RoboDK station: PRBE_Operateur_v2.rdk

Station PRBE_Operateur_v2 (saved by RoboDK 6.0.4). Poses are relative to the parent item; angles as X-Y-Z fixed-axis rotations.
  - object Manikin_1 at (0, 0, 0) mm, geometry from Manikin_1.STEP
  - frame Human_Base at (0, 958, 0) mm
    - item type 7 Manikin_1-bassin
    - item type 7 Manikin_1-torso
    - item type 7 Manikin_1-tete
    - frame hipL_abduction at (63.26, -78.51, -37.42) mm
      - frame hipL_flexion at (0, 0, 0) mm
        - frame hipL_rotation at (0, 0, 0) mm
          - item type 7 Manikin_1-cuisse_g
          - frame kneeL_flexion at (67.44, -393.44, -12.97) mm
            - item type 7 Manikin_1-tibia_g
            - frame ankleL_flexion at (42.46, -394.54, 0) mm
              - item type 7 Manikin_1-pied_g
    - frame shoulderL_abduction at (206.4, 423.68, 12.96) mm, rotated rx 0 ry 0 rz -42 deg
      - frame shoulderL_flexion at (0, 0, 0) mm
        - frame shoulderL_rotation at (0, 0, 0) mm
          - item type 7 Manikin_1-bras_g
          - frame elbowL_flexion at (155.8, -191.9, 27.9) mm
            - item type 7 Manikin_1-avant_bras_g
            - frame wristL_flexion at (148.7, -146.81, 80.89) mm
              - frame wristL_deviation at (0, 0, 0) mm
                - item type 7 Manikin_1-main_g
    - frame hipR_abduction at (-70.11, -75.34, -37.06) mm
      - frame hipR_flexion at (0, 0, 0) mm
        - frame hipR_rotation at (0, 0, 0) mm
          - item type 7 Manikin_1-cuisse_d
          - frame kneeR_flexion at (-86.5, -385.51, -37.91) mm
            - item type 7 Manikin_1-tibia_d_1
            - item type 7 Manikin_1-tibia_d_2
            - frame ankleR_flexion at (-60.5, -382.31, -26.03) mm
              - item type 7 Manikin_1-pied_d_1
              - item type 7 Manikin_1-pied_d_2
    - frame shoulderR_abduction at (-133.98, 420.49, -26.02) mm
      - frame shoulderR_flexion at (0, 0, 0) mm
        - frame shoulderR_rotation at (0, 0, 0) mm
          - item type 7 Manikin_1-bras_d
          - frame elbowR_flexion at (-80.76, -228.86, 52.14) mm
            - item type 7 Manikin_1-avant_bras_d
            - frame wristR_flexion at (-76.34, -195.54, 87.27) mm
              - frame wristR_deviation at (0, 0, 0) mm
                - item type 7 Manikin_1-main_d
  - Python program Mouvement_v2 (listed below)
  - Python program Marche_Militaire (listed below)
  - Python program Marche_Avant (listed below)

--- Python program Mouvement_v2 ---
# -*- coding: utf-8 -*-
"""
Mouvement_v2.py — MODELE pour piloter l'operateur v2 (22 DDL).

A LANCER DANS ROBODK (clic droit > Run) depuis la station PRBE_Operateur_v2,
operateur en pose NEUTRE (le script capture le repos au demarrage).

PRINCIPE :
  - chaque DDL = un repere nomme (ex: "hipR_flexion") qui tourne sur UN axe.
  - bouge("nom_du_ddl", angle_en_degres) tourne ce DDL depuis le repos.
  - les angles sont automatiquement borns aux limites du corps humain.
"""
from robolink import Robolink
from robodk.robomath import rotx, roty, rotz
import math
import time

RDK = Robolink()

# ---- Les 22 DDL : nom -> (axe, limite_basse_deg, limite_haute_deg) ----
DDL = {
    # JAMBE DROITE (5)
    "hipR_abduction": ("z", -45, 30),   "hipR_flexion": ("x", -120, 15),  "hipR_rotation": ("y", -45, 45),
    "kneeR_flexion":  ("x", 0, 135),    "ankleR_flexion": ("x", -30, 50),
    # JAMBE GAUCHE (5)
    "hipL_abduction": ("z", -30, 45),   "hipL_flexion": ("x", -120, 15),  "hipL_rotation": ("y", -45, 45),
    "kneeL_flexion":  ("x", 0, 135),    "ankleL_flexion": ("x", -30, 50),
    # BRAS DROIT (6)
    "shoulderR_abduction": ("z", -135, 90), "shoulderR_flexion": ("x", -90, 90), "shoulderR_rotation": ("y", -45, 180),
    "elbowR_flexion": ("x", 0, 145),
    "wristR_flexion": ("x", -50, 60),   "wristR_deviation": ("z", -30, 20),
    # BRAS GAUCHE (6)
    "shoulderL_abduction": ("z", -90, 135), "shoulderL_flexion": ("x", -90, 90), "shoulderL_rotation": ("y", -45, 180),
    "elbowL_flexion": ("x", 0, 145),
    "wristL_flexion": ("x", -50, 60),   "wristL_deviation": ("z", -30, 20),
}

ROT = {"x": rotx, "y": roty, "z": rotz}
F = {nom: RDK.Item(nom) for nom in DDL}            # les reperes
REST = {nom: F[nom].Pose() for nom in DDL}         # pose neutre (capturee au demarrage)


def bouge(nom, deg):
    """Tourne un DDL de `deg` degres depuis le repos (born aux limites)."""
    axe, lo, hi = DDL[nom]
    deg = max(lo, min(hi, deg))                    # ne depasse pas le corps humain
    F[nom].setPose(REST[nom] * ROT[axe](math.radians(deg)))


def neutre():
    """Remet tout l'operateur droit."""
    for nom in DDL:
        F[nom].setPose(REST[nom])


# =======================================================================
# TON CODE ICI. Exemples :
# =======================================================================

# --- EXEMPLE 1 : une pose (lever le bras droit + plier le coude) ---
bouge("shoulderR_flexion", -70)   # bras droit vers l'avant
bouge("elbowR_flexion", 90)       # coude plie
RDK.Render(True)
time.sleep(1)

# --- EXEMPLE 2 : une petite animation (le bras qui salue) ---
neutre()
bouge("shoulderR_abduction", 80)  # bras leve sur le cote
for i in range(6):
    RDK.Render(False)
    bouge("elbowR_flexion", 30 + 40 * (i % 2))   # avant-bras qui va et vient
    RDK.Render(True)
    time.sleep(0.3)

neutre()
RDK.Render(True)
print("Fini.")

--- Python program Marche_Militaire ---
# -*- coding: utf-8 -*-
"""
Marche_Militaire.py — L'operateur marque le pas (marche militaire sur place).

A LANCER DANS ROBODK (clic droit > Run) depuis la station avec le rig 22 DDL,
operateur en pose NEUTRE (le script capture le repos au demarrage).

Principe de la marche militaire :
  - genoux qui montent haut, alternes
  - bras RAIDES (coude quasi tendu) qui balancent en OPPOSITION des jambes
  - buste droit (il est fige, parfait pour un militaire)

Regle les amplitudes/vitesse dans la section REGLAGES.
"""
from robolink import Robolink
from robodk.robomath import rotx, roty, rotz
import math
import time

RDK = Robolink()

# ---- Les 22 DDL : nom -> (axe, limite_basse_deg, limite_haute_deg) ----
DDL = {
    # JAMBE DROITE (5)
    "hipR_abduction": ("z", -45, 30),   "hipR_flexion": ("x", -120, 15),  "hipR_rotation": ("y", -45, 45),
    "kneeR_flexion":  ("x", 0, 135),    "ankleR_flexion": ("x", -30, 50),
    # JAMBE GAUCHE (5)
    "hipL_abduction": ("z", -30, 45),   "hipL_flexion": ("x", -120, 15),  "hipL_rotation": ("y", -45, 45),
    "kneeL_flexion":  ("x", 0, 135),    "ankleL_flexion": ("x", -30, 50),
    # BRAS DROIT (6)
    "shoulderR_abduction": ("z", -135, 90), "shoulderR_flexion": ("x", -90, 90), "shoulderR_rotation": ("y", -45, 180),
    "elbowR_flexion": ("x", 0, 145),
    "wristR_flexion": ("x", -50, 60),   "wristR_deviation": ("z", -30, 20),
    # BRAS GAUCHE (6)
    "shoulderL_abduction": ("z", -90, 135), "shoulderL_flexion": ("x", -90, 90), "shoulderL_rotation": ("y", -45, 180),
    "elbowL_flexion": ("x", 0, 145),
    "wristL_flexion": ("x", -50, 60),   "wristL_deviation": ("z", -30, 20),
}

ROT = {"x": rotx, "y": roty, "z": rotz}
F = {nom: RDK.Item(nom) for nom in DDL}            # les reperes
REST = {nom: F[nom].Pose() for nom in DDL}         # pose neutre (capturee au demarrage)


def bouge(nom, deg):
    """Tourne un DDL de `deg` degres depuis le repos (borne aux limites)."""
    axe, lo, hi = DDL[nom]
    deg = max(lo, min(hi, deg))
    F[nom].setPose(REST[nom] * ROT[axe](math.radians(deg)))


def neutre():
    """Remet tout l'operateur droit."""
    for nom in DDL:
        F[nom].setPose(REST[nom])


# =======================================================================
# REGLAGES de la marche militaire
# =======================================================================
HANCHE = 55      # levee de cuisse (deg) — genou haut
GENOU = 65       # pliage du genou quand la jambe monte (deg)
CHEVILLE = 15    # pointe de pied quand la jambe est levee (deg)
BRAS_AV = -45    # bras vers l'AVANT (deg, negatif = devant)
BRAS_ARR = 20    # bras vers l'ARRIERE (deg)
COUDE = 8        # coude quasi tendu = bras raide militaire
NB_PAS = 8       # nombre de pas au total
IMAGES_PAR_PAS = 12   # fluidite (images par pas)
DT = 0.04        # pause entre images (s) — plus petit = plus rapide


def pose_marche(ph):
    """Pose complete de la marche pour une phase `ph` (radians).
       Jambe droite levee sur [0, pi], jambe gauche sur [pi, 2pi]."""
    s = math.sin(ph)
    lift_d = max(0.0, s)     # jambe droite qui monte
    lift_g = max(0.0, -s)    # jambe gauche qui monte

    # jambes : genou haut + pointe de pied
    bouge("hipR_flexion", -HANCHE * lift_d)
    bouge("kneeR_flexion", GENOU * lift_d)
    bouge("ankleR_flexion", CHEVILLE * lift_d)
    bouge("hipL_flexion", -HANCHE * lift_g)
    bouge("kneeL_flexion", GENOU * lift_g)
    bouge("ankleL_flexion", CHEVILLE * lift_g)

    # bras raides, en opposition : bras droit devant quand jambe gauche monte
    u_d = (1.0 - s) / 2.0    # 0 = bras D derriere, 1 = bras D devant
    u_g = (1.0 + s) / 2.0
    bouge("shoulderR_flexion", BRAS_ARR + (BRAS_AV - BRAS_ARR) * u_d)
    bouge("shoulderL_flexion", BRAS_ARR + (BRAS_AV - BRAS_ARR) * u_g)
    bouge("elbowR_flexion", COUDE)
    bouge("elbowL_flexion", COUDE)


def marche(nb_pas=NB_PAS, images_par_pas=IMAGES_PAR_PAS, dt=DT):
    """Anime la marche militaire sur place."""
    for i in range(nb_pas * images_par_pas + 1):
        ph = math.pi * i / images_par_pas      # 1 pas = une demi-periode
        RDK.Render(False)
        pose_marche(ph)
        RDK.Render(True)
        time.sleep(dt)
    neutre()
    RDK.Render(True)


if __name__ == "__main__":
    print("Marche militaire : {} pas...".format(NB_PAS))
    marche()
    print("Repos !")

--- Python program Marche_Avant ---
# -*- coding: utf-8 -*-
"""
Marche_Avant.py — L'operateur marche TOUT DROIT devant lui (marche naturelle).

A LANCER DANS ROBODK (clic droit > Run) depuis la station avec le rig 22 DDL,
operateur au repos / garde-a-vous (le script capture le repos au demarrage).

Principe :
  - hanches qui balancent avant/arriere, genou qui se plie pendant le balance
  - bras souples en opposition des jambes (coude legerement plie)
  - le CORPS AVANCE a la vitesse des pas (longueur de pas calculee depuis
    l'amplitude de hanche) -> pas de glisse visible
  - il marche vers SON regard (+Z monde). A la fin, il REVIENT au centre
    (position d'origine de Human_Base).

Regle les amplitudes/vitesse dans la section REGLAGES.
"""
from robolink import Robolink
from robodk.robomath import rotx, roty, rotz, transl
import math
import time

RDK = Robolink()

# ---- Les 22 DDL : nom -> (axe, limite_basse_deg, limite_haute_deg) ----
DDL = {
    # JAMBE DROITE (5)
    "hipR_abduction": ("z", -45, 30),   "hipR_flexion": ("x", -120, 15),  "hipR_rotation": ("y", -45, 45),
    "kneeR_flexion":  ("x", 0, 135),    "ankleR_flexion": ("x", -30, 50),
    # JAMBE GAUCHE (5)
    "hipL_abduction": ("z", -30, 45),   "hipL_flexion": ("x", -120, 15),  "hipL_rotation": ("y", -45, 45),
    "kneeL_flexion":  ("x", 0, 135),    "ankleL_flexion": ("x", -30, 50),
    # BRAS DROIT (6)
    "shoulderR_abduction": ("z", -135, 90), "shoulderR_flexion": ("x", -90, 90), "shoulderR_rotation": ("y", -45, 180),
    "elbowR_flexion": ("x", 0, 145),
    "wristR_flexion": ("x", -50, 60),   "wristR_deviation": ("z", -30, 20),
    # BRAS GAUCHE (6)
    "shoulderL_abduction": ("z", -90, 135), "shoulderL_flexion": ("x", -90, 90), "shoulderL_rotation": ("y", -45, 180),
    "elbowL_flexion": ("x", 0, 145),
    "wristL_flexion": ("x", -50, 60),   "wristL_deviation": ("z", -30, 20),
}

ROT = {"x": rotx, "y": roty, "z": rotz}
F = {nom: RDK.Item(nom) for nom in DDL}            # les reperes
REST = {nom: F[nom].Pose() for nom in DDL}         # pose de repos (capturee au demarrage)
BASE = RDK.Item("Human_Base")
BASE_REST = BASE.Pose()                            # position de depart du corps
HOME = transl(0, 958, 0)                           # position d'origine (au centre, 1er repere)


def bouge(nom, deg):
    """Tourne un DDL de `deg` degres depuis le repos (borne aux limites)."""
    axe, lo, hi = DDL[nom]
    deg = max(lo, min(hi, deg))
    F[nom].setPose(REST[nom] * ROT[axe](math.radians(deg)))


def neutre():
    """Remet les articulations au repos (le corps reste ou il est)."""
    for nom in DDL:
        F[nom].setPose(REST[nom])


# =======================================================================
# REGLAGES de la marche
# =======================================================================
HANCHE_AV = 30    # jambe vers l'avant (deg)
HANCHE_ARR = 12   # jambe vers l'arriere (deg)
GENOU = 50        # pliage du genou pendant le balance (deg)
CHEVILLE = 8      # pointe de pied relevee pendant le balance (deg)
BRAS_AV = 25      # bras vers l'avant (deg)
BRAS_ARR = 15     # bras vers l'arriere (deg)
COUDE = 20        # coude legerement plie (marche naturelle)
NB_PAS = 8        # nombre de pas
IMAGES_PAR_PAS = 14   # fluidite
DT = 0.04         # pause entre images (s)

LONGUEUR_JAMBE = 790.0   # hanche -> cheville (mm, mesure sur le modele)
SENS = +1                # +1 = devant lui (+Z monde). Mets -1 pour marche arriere.

# longueur d'un pas deduite du balancement de hanche (pour avancer sans glisser)
LONGUEUR_PAS = LONGUEUR_JAMBE * (math.sin(math.radians(HANCHE_AV)) + math.sin(math.radians(HANCHE_ARR)))


def pose_pas(ph):
    """Pose de marche pour une phase `ph` (radians). Jambe droite devant sur [0, pi]."""
    s = math.sin(ph)
    # hanches : avant = negatif (amplitude asymetrique avant/arriere)
    a = (HANCHE_AV + HANCHE_ARR) / 2.0
    c = (HANCHE_AV - HANCHE_ARR) / 2.0
    bouge("hipR_flexion", -(a * s + c))
    bouge("hipL_flexion", -(a * -s + c))
    # genou plie pendant le balance (jambe qui revient vers l'avant)
    bouge("kneeR_flexion", GENOU * max(0.0, math.cos(ph)))
    bouge("kneeL_flexion", GENOU * max(0.0, -math.cos(ph)))
    # pointe de pied relevee pendant le balance (pour ne pas racler le sol)
    bouge("ankleR_flexion", -CHEVILLE * max(0.0, math.cos(ph)))
    bouge("ankleL_flexion", -CHEVILLE * max(0.0, -math.cos(ph)))
    # bras en opposition, coude souple
    sa = (BRAS_AV + BRAS_ARR) / 2.0
    sc = (BRAS_ARR - BRAS_AV) / 2.0
    bouge("shoulderR_flexion", sa * s + sc)
    bouge("shoulderL_flexion", -sa * s + sc)
    bouge("elbowR_flexion", COUDE)
    bouge("elbowL_flexion", COUDE)


def avance(dist):
    """Place le corps a `dist` mm devant sa position de depart."""
    BASE.setPose(BASE_REST * transl(0, 0, SENS * dist))


def marche(nb_pas=NB_PAS, images_par_pas=IMAGES_PAR_PAS, dt=DT):
    """Anime la marche en avant, puis remet l'operateur au centre (HOME)."""
    for i in range(nb_pas * images_par_pas + 1):
        ph = math.pi * i / images_par_pas      # 1 pas = une demi-periode
        RDK.Render(False)
        pose_pas(ph)
        avance(LONGUEUR_PAS * ph / math.pi)
        RDK.Render(True)
        time.sleep(dt)
    # fin : repos + retour a la position initiale, au centre
    RDK.Render(False)
    neutre()
    BASE.setPose(HOME)
    RDK.Render(True)


if __name__ == "__main__":
    d_tot = LONGUEUR_PAS * NB_PAS / 1000.0
    print("Marche avant : {} pas (~{:.1f} m)...".format(NB_PAS, d_tot))
    marche()
    print("Arrive !")
